(* IEC 61131-3 sources: plc-vscode/tests/st/all/rusty/tests/lit/single/functions, 8 files *)

(* ---- call_with_array_access_on_result.st ---- *)
// RUN: (%COMPILE %s && %RUN) | %CHECK %s

FUNCTION foo: ARRAY[1..5] OF DINT
    foo := [5, 4, 3, 2, 1];
END_FUNCTION

FUNCTION alwaysOne: DINT
    alwaysOne := 1;
END_FUNCTION

FUNCTION main
    VAR
        value: DINT;
        one: DINT := 1;
        two: DINT := 2;
    END_VAR

    // CHECK: 5
    value := foo()[1];
    printf('%d$N', value);

    // CHECK: 3
    value := foo()[1 + 2];
    printf('%d$N', value);

    // CHECK: 5
    value := foo()[one];
    printf('%d$N', value);

    // CHECK: 3
    value := foo()[one + two];
    printf('%d$N', value);

    // CHECK: 5
    value := foo()[alwaysOne()];
    printf('%d$N', value);
END_FUNCTION

(* ---- default_params.st ---- *)
// RUN: (%COMPILE %s && %RUN) | %CHECK %s
FUNCTION func : int
  VAR_INPUT
    in : INT := 42;
  END_VAR
  func := in;
END_FUNCTION

FUNCTION main : DINT

    PRINTF('func complete:%d$N', func(13)); //CHECK: func complete:13
    PRINTF('func incomplete:%d$N', func()); //CHECK: func incomplete:42

END_FUNCTION

(* ---- function_output_should_be_cast_if_needed.st ---- *)
// RUN: (%COMPILE %s && %RUN) | %CHECK %s
FUNCTION outputCastIntToReal : INT
    VAR_OUTPUT
        result : REAL;
    END_VAR

    result := 42.0;
END_FUNCTION

FUNCTION outputNoCastInt : INT
    VAR_OUTPUT
        result : INT;
    END_VAR

    result := 52;
END_FUNCTION

FUNCTION outputCastRealToInt : INT
    VAR_OUTPUT
        result : INT;
    END_VAR

    result := 62;
END_FUNCTION

FUNCTION outputNoCastReal : INT
    VAR_OUTPUT
        result : REAL;
    END_VAR

    result := 72.0;
END_FUNCTION

FUNCTION main
    VAR
        i1 : INT;
        i2 : INT;
        r1 : REAL;
        r2 : REAL;
    END_VAR

    i1 := 31;
    i2 := 32;
    r1 := 33;
    r2 := 34;

    // ----------------- //
    // -- INT to REAL -- //

    outputCastIntToReal(
        result => i1
    );

    // CHECK: 42
    PRINTF('%d$N', i1);

    // ---------------- //
    // -- INT to INT -- //

    outputNoCastInt(
        result => i2
    );

    // CHECK: 52
    PRINTF('%d$N', i2);

    // ----------------- //
    // -- REAL to INT -- //

    outputCastRealToInt(
        result => r1
    );

    // CHECK: 62.0
    PRINTF('%.1f$N', r1);

    // ------------------ //
    // -- REAL to REAL -- //

    outputNoCastReal(
        result => r2
    );

    // CHECK: 72.0
    PRINTF('%.1f$N', r2);
END_FUNCTION

(* ---- function_parameter_with_bit_access.st ---- *)
// RUN: (%COMPILE %s && %RUN) | %CHECK %s
FUNCTION FLIP
    VAR_INPUT
        in: BYTE;
    END_VAR
    VAR_OUTPUT
        out : BYTE;
    END_VAR
    out := NOT(in);
END_FUNCTION

FUNCTION main
    VAR
        wordVar : WORD;
    END_VAR

    wordVar := 0;
    FLIP(2#01010101, wordVar.%b0);

    // CHECK: wordVar=170
    PRINTF('wordVar=%d$N', wordVar);
END_FUNCTION

(* ---- function_parameter_with_bit_access_named_params.st ---- *)
// RUN: (%COMPILE %s && %RUN) | %CHECK %s
FUNCTION FLIP
    VAR_INPUT
        in: BYTE;
    END_VAR
    VAR_OUTPUT
        out : BYTE;
    END_VAR
    out := NOT(in);
END_FUNCTION

FUNCTION main
    VAR
        wordVar : WORD;
    END_VAR

    wordVar := 0;
    FLIP(in := 2#01010101, out => wordVar.%b0);

    // CHECK: wordVar=170
    PRINTF('wordVar=%d$N', wordVar);
END_FUNCTION

(* ---- function_block_output_should_be_cast_if_needed.st ---- *)
// RUN: (%COMPILE %s && %RUN) | %CHECK %s
FUNCTION_BLOCK outputCastIntToReal_fb
    VAR_OUTPUT
        result : REAL;
    END_VAR

    result := 42.0;
END_FUNCTION_BLOCK

FUNCTION_BLOCK outputNoCastInt_fb
    VAR_OUTPUT
        result : INT;
    END_VAR

    result := 52;
END_FUNCTION_BLOCK

FUNCTION_BLOCK outputCastRealToInt_fb
    VAR_OUTPUT
        result : INT;
    END_VAR

    result := 62;
END_FUNCTION_BLOCK

FUNCTION_BLOCK outputNoCastReal_fb
    VAR_OUTPUT
        result : REAL;
    END_VAR

    result := 72.0;
END_FUNCTION_BLOCK

FUNCTION main
    VAR
        outputCastIntToReal : outputCastIntToReal_fb;
        outputNoCastInt : outputNoCastInt_fb;
        outputCastRealToInt : outputCastRealToInt_fb;
        outputNoCastReal : outputNoCastReal_fb;

        i1 : INT;
        i2 : INT;
        r1 : REAL;
        r2 : REAL;
    END_VAR

    i1 := 31;
    i2 := 32;
    r1 := 33;
    r2 := 34;

    // ----------------- //
    // -- INT to REAL -- //

    outputCastIntToReal(
        result => i1
    );

    // CHECK: 42
    PRINTF('%d$N', i1);

    // ---------------- //
    // -- INT to INT -- //

    outputNoCastInt(
        result => i2
    );

    // CHECK: 52
    PRINTF('%d$N', i2);

    // ----------------- //
    // -- REAL to INT -- //

    outputCastRealToInt(
        result => r1
    );

    // CHECK: 62.0
    PRINTF('%.1f$N', r1);

    // ------------------ //
    // -- REAL to REAL -- //

    outputNoCastReal(
        result => r2
    );

    // CHECK: 72.0
    PRINTF('%.1f$N', r2);
END_FUNCTION

(* ---- function_output_to_bit_direct_access.st ---- *)
// RUN: (%COMPILE %s && %RUN) | %CHECK %s

// Regression test for https://github.com/PLC-lang/rusty/issues/1239
// `fun(out => bar.4)` and `myFb(out => bar.4)` previously generated IR that
// computed the bit address but never stored the function's output back into
// the underlying integer.
FUNCTION fun
    VAR_OUTPUT
        foo : BOOL;
    END_VAR
    foo := TRUE;
END_FUNCTION

FUNCTION_BLOCK fb
    VAR_OUTPUT
        foo : BOOL;
    END_VAR
    foo := TRUE;
END_FUNCTION_BLOCK

FUNCTION main : DINT
    VAR
        bar  : DINT;
        myFb : fb;
    END_VAR

    bar := 0;
    fun(foo => bar.4);
    PRINTF('after_fun=%d$N', bar);
    // CHECK: after_fun=16

    bar := 0;
    myFb(foo => bar.4);
    PRINTF('after_fb=%d$N', bar);
    // CHECK: after_fb=16

    // Non-zero seed: anchors that bits 0–3 are *preserved* when the FB output
    // writes bit 4. A regression that clobbered the integer (e.g. wrote a full
    // word instead of just the bit) would surface here as 16 instead of 17.
    bar := 1;
    myFb(foo => bar.4);
    PRINTF('after_fb_seeded=%d$N', bar);
    // CHECK: after_fb_seeded=17
END_FUNCTION

(* ---- segmented_variable_blocks_with_implicit_arguments_call.st ---- *)
// RUN: (%COMPILE %s && %RUN) | %CHECK %s

FUNCTION_BLOCK foo
    VAR
        placeholder_one: DINT;
    END_VAR

    VAR_INPUT
        a, b: DINT;
    END_VAR

    VAR
        placeholder_two: DINT;
    END_VAR

    VAR_OUTPUT
        c: DINT;
    END_VAR

    c := a + b;
END_FUNCTION_BLOCK

FUNCTION main
    VAR
        foo: foo;
        local_a, local_b, local_c: DINT := 2;
    END_VAR

    foo(local_a, local_b, local_c);
    printf('%d$N', local_c); // CHECK: 4
END_FUNCTION
